(* IEC 61131-3 sources: NachHouse_TST/ROOM_API_PILOT/room_api_pilot, 11 files *)

(* ---- 02_TYPES.ST ---- *)
(*
   ROOM_API_PILOT - d�tov� typy logick�ho API a prenosov�ho protokolu.
   Koment�re opisuj� v�znam pre PLC aj klienta; nejde o re�lnu domov� automatiz�ciu.
*)

TYPE
   NH_API_INFO : STRUCT
    	ApiVersion		: UINT;          (* Verzia verejn�ho API kontraktu. ENG *)
		ApiVarNext		: UINT;          (* Adresa v pam�ti PLC, kde sa nach�dza za�iatok �al��ch premenn�ch API. ENG *)
		ApiVarSize		: UDINT;          (* Ve�kos� v bajtoch, ktor� zaber� v pam�ti PLC. ENG *)
		ApiBussy			: BOOL;          (* TRUE znamen�, �e PLC je zanepr�znene spracovan�m pr�kazu. ENG *)
   END_STRUCT

   NH_LOG_INFO : STRUCT
		BufferBegin		: UDINT;          (* Adresa v pam�ti PLC, kde sa nach�dza za�iatok logovacieho bufferu. ENG *)
		BufferEnd		: UDINT;          (* Adresa v pamti PLC, kde sa nachdza zaiatok logovacieho bufferu. ENG *)
		BufferNext		: UDINT;          (* Adresa v pamti PLC, kde sa nachdza zaiatokalch premennch API. ENG *)
		BufferSize		: UDINT;          (* Vekos v bajtoch, ktor zaber v pamti PLC. ENG *)
   END_STRUCT

END_TYPE

TYPE
    NH_API_DIFF_HEAD : STRUCT                    (* Header pre diff udajov, Sizeof = 40B *)
        StructID        : UINT := 1;          		(* Cislo struktury zaslatych udajov - parser  *)
        Name            : STRING[21] := 'T_ROOM_STATE';   (* What scheme used for parser. StructID = 1 = T_ROOM_STATE*)
        Records         : INT := 2;          		(* Pocet zaslatych zaznamov T_ROOM_STATE *)
        RecSize         : UDINT := 21;      			(* Size of 1. T_ROOM_STATE*)
        MessageSize     : UDINT := 42;      			(* Len Doplnujuce info Records * RecSize := 2*21=42B *)
        HeadIndex       : UINT := 0;						(* index tohto headera ApiVarsPublic[0], koniec ApiVarsPublic[0] + 40B = ApiVarsPublic[3] *)
        BeginIndex      : UINT := 4;          		(* kde zacinaju data struktury = 1.veta ApiVarsPublic[4] *)
        EndIndex        : UINT := 8;          		(* kde koncia data ApiVarsPublic[8] .. len informacne, lebo nemusi byt zaplnenychcelych 4B DWORD *)
	END_STRUCT

	T_ROOM_STATE : STRUCT
      RoomId          : UDINT; (* V?zba stavov?ho z?znamu na stabiln? ID v konfigur?cii. ENG *)
    	Temperature     : REAL;  (* Zobrazovan? testovacia teplota v stup?och Celzia. ENG *)
    	Humidity        : REAL;  (* Zobrazovan? testovacia relat?vna vlhkos? v percent?ch. ENG *)
    	Presence        : BOOL;  (* Testovac? pr?znak pr?tomnosti ovplyv?uj?ci pozadie karty. ENG *)
    	DayPhase        : UINT;  (* K?d dennej f?zy API_DAY_PHASE_* pre existuj?cu ikonu. ENG *)
    	CategoryMask    : DWORD; (* Bitov? maska kateg?ri?, ktor?ch ikony sa maj? zobrazi?. ENG *)
    	AlarmLevel      : USINT; (* Vizu?lna ?rove? API_ALARM_*; nesp???a re?lny alarm. ENG *)
    	Online          : BOOL;  (* Dostupnos? d?t miestnosti pre klienta. ENG *)
	END_STRUCT
END_TYPE
TYPE
   NH_API_DIFF_HEAD : STRUCT                    (* Header pre diff udajov, Sizeof = 40B *)
		StructID		: UINT := 1;          		(* Cislo struktury zaslatych udajov - parser  *)
		Name			: STRING[21] := 'T_ROOM_STATE';   (* What scheme used for parser. StructID = 1 = T_ROOM_STATE*)
		Records			: INT := 2;          		(* Pocet zaslatych zaznamov T_ROOM_STATE *)
		RecSize			: UDINT := 21;      			(* Size of 1. T_ROOM_STATE*)
		MessageSize		: UDINT := 42;      			(* Len Doplnujuce info Records * RecSize := 2*21=42B *)
         HeadIndex      : UINT := 0;						(* index tohto headera ApiVarsPublic[0], koniec ApiVarsPublic[0] + 40B = ApiVarsPublic[3] *)
		BeginIndex		: UINT := 4;          		(* kde zacinaju data struktury = 1.veta ApiVarsPublic[4] *)
		EndIndex		: UINT := 8;          		(* kde koncia data ApiVarsPublic[8] .. len informacne, lebo nemusi byt zaplnenychcelych 4B DWORD *)
	END_STRUCT

	T_ROOM_STATE : STRUCT
   	    RoomId          : UDINT; (* V�zba stavov�ho z�znamu na stabiln� ID v konfigur�cii. ENG *)
    	Temperature     : REAL;  (* Zobrazovan� testovacia teplota v stup�och Celzia. ENG *)
    	Humidity        : REAL;  (* Zobrazovan� testovacia relat�vna vlhkos� v percent�ch. ENG *)
    	Presence        : BOOL;  (* Testovac� pr�znak pr�tomnosti ovplyv�uj�ci pozadie karty. ENG *)
    	DayPhase        : UINT;  (* K�d dennej f�zy API_DAY_PHASE_* pre existuj�cu ikonu. ENG *)
    	CategoryMask    : DWORD; (* Bitov� maska kateg�ri�, ktor�ch ikony sa maj� zobrazi�. ENG *)
    	AlarmLevel      : USINT; (* Vizu�lna �rove� API_ALARM_*; nesp���a re�lny alarm. ENG *)
    	Online          : BOOL;  (* Dostupnos� d�t miestnosti pre klienta. ENG *)
	END_STRUCT
END_TYPE

(* V�sledok vykonania jedn�ho klientsk�ho pr�kazu. *)
TYPE
T_API_COMMAND_RESULT : STRUCT
    ClientId       : STRING[36]; (* Identifik�tor klienta, ktor�mu patr� v�sledok. ENG *)
    RequestId      : UDINT;      (* Identifik�tor po�iadavky pridelen� klientom. ENG *)
    Result         : USINT;      (* ��seln� n�vratov� k�d API_RESULT_*. ENG *)
    Message        : STRING[80]; (* Kr�tky slovensk� text v�sledku ur�en� pre log a testovanie. *)
    ConfigRevision : UDINT;      (* Rev�zia konfigur�cie platn� po spracovan� pr�kazu. ENG *)
    StateRevision  : UDINT;      (* Rev�zia stavov�ch �dajov platn� po spracovan� pr�kazu. ENG *)
END_STRUCT
END_TYPE

(* Z�kladn� inform�cie o API a jeho aktu�lnych rev�zi�ch. *)
TYPE T_API_INFO :
STRUCT
    ApiVersion        : STRING[32];          (* Verzia verejn�ho API kontraktu. ENG *)
    ConfigRevision    : UDINT;               (* Aktu�lna rev�zia konfigur�cie miestnost�. ENG *)
    StateRevision     : UDINT;               (* Aktu�lna rev�zia dynamick�ch stavov miestnost�. ENG *)
    MaxRooms          : USINT;               (* Najvy��� po�et miestnost� podporovan� PLC. ENG *)
    LastCommandResult : T_API_COMMAND_RESULT; (* Posledn� v�sledok pr�kazu, dostupn� aj po obnoven� klienta. ENG *)
END_STRUCT
END_TYPE

(* Konfigura�n� �daje jednej miestnosti. *)
TYPE T_ROOM_CONFIG :
STRUCT
    Used        : BOOL;       (* TRUE znamen�, �e je t�to poz�cia po�a obsaden� miestnos�ou. ENG *)
    RoomId      : UDINT;      (* Stabiln� a jedine�n� identifik�tor miestnosti; hodnota 0 je neplatn�. ENG *)
    Name        : STRING[64]; (* Hlavn� n�zov miestnosti zobrazen� na karte. ENG *)
    ProjectName : STRING[64]; (* Doplnkov� n�zov zobrazen� pod hlavn�m n�zvom. ENG *)
    IconId      : UINT;       (* Identifik�tor ikony pou��vanej frozen browserom. ENG *)
    SortDefault : UINT;       (* Predvolen� poradie iba pri prvom na��tan� klienta. ENG *)
END_STRUCT
END_TYPE

(* �pln� konfigura�n� snapshot v�etk�ch poz�ci� miestnost�. *)
TYPE T_API_CONFIG :
STRUCT
    Rooms : ARRAY[1..40] OF T_ROOM_CONFIG; (* Pevn� pole najviac 40 konfigura�n�ch z�znamov. ENG *)
END_STRUCT
END_TYPE

(* Ru�ne nastavovan� pilotn� stav jednej miestnosti. *)

(* �pln� stavov� snapshot v�etk�ch poz�ci� miestnost�. *)
TYPE T_API_STATE :
STRUCT
    Rooms : ARRAY[1..40] OF T_ROOM_STATE; (* Pevn� pole najviac 40 stavov�ch z�znamov. ENG *)
END_STRUCT
END_TYPE

(* Po�iadavka klienta na pridanie, zmazanie, kop�rovanie alebo �pravu miestnosti. *)
TYPE T_API_COMMAND_ROOM :
STRUCT
    ClientId     : STRING[36]; (* Identifik�tor klienta odosielaj�ceho pr�kaz. ENG *)
    RequestId    : UDINT;      (* Nenulov� identifik�tor po�iadavky pre p�rovanie a opakovanie. ENG *)
    Action       : USINT;      (* Po�adovan� akcia ur�en� kon�tantou API_ACTION_*. ENG *)
    RoomId       : UDINT;      (* Cie�ov� stabiln� ID miestnosti. ENG *)
    SourceRoomId : UDINT;      (* Zdrojov� ID pou�it� iba pri kop�rovan� miestnosti. ENG *)
    Name         : STRING[64]; (* Nov� alebo upraven� hlavn� n�zov miestnosti. ENG *)
    ProjectName  : STRING[64]; (* Nov� alebo upraven� doplnkov� n�zov miestnosti. ENG *)
END_STRUCT
END_TYPE

(* Jedna polo�ka konfigura�n�ho diffu. *)
TYPE T_API_CONFIG_CHANGE :
STRUCT
    Valid     : BOOL;          (* TRUE znamen�, �e polo�ka obsahuje platn� zmenu. ENG *)
    Operation : USINT;         (* Druh zmeny API_DIFF_UPSERT alebo API_DIFF_DELETE. ENG *)
    RoomId    : UDINT;         (* Stabiln� ID zmenenej alebo odstr�nenej miestnosti. ENG *)
    Room      : T_ROOM_CONFIG; (* �pln� nov� z�znam pri UPSERT; pri DELETE je vy�isten�. ENG *)
END_STRUCT
END_TYPE

(* Jedna polo�ka stavov�ho diffu. *)
TYPE T_API_STATE_CHANGE :
STRUCT
    Valid     : BOOL;         (* TRUE znamen�, �e polo�ka obsahuje platn� zmenu. ENG *)
    Operation : USINT;        (* Druh zmeny API_DIFF_UPSERT alebo API_DIFF_DELETE. ENG *)
    RoomId    : UDINT;        (* Stabiln� ID zmenen�ho alebo odstr�nen�ho stavu. ENG *)
    Room      : T_ROOM_STATE; (* �pln� nov� stav pri UPSERT; pri DELETE je vy�isten�. ENG *)
END_STRUCT
END_TYPE

(* Jeden rev�zny r�mec zmien konfigur�cie. *)
TYPE T_API_CONFIG_DIFF :
STRUCT
    Valid        : BOOL;  (* TRUE znamen�, �e hlavi�ka a obsah r�mca s� pripraven�. ENG *)
    FromRevision : UDINT; (* Rev�zia, na ktor� tento r�mec priamo nadv�zuje. ENG *)
    ToRevision   : UDINT; (* Rev�zia po aplikovan� v�etk�ch zmien z r�mca. ENG *)
    FullRequired : BOOL;  (* TRUE prikazuje klientovi na��ta� cel� snapshot. ENG *)
    ChangeCount  : USINT; (* Po�et platn�ch polo�iek na za�iatku po�a Changes. ENG *)
    Changes      : ARRAY[1..40] OF T_API_CONFIG_CHANGE; (* Zmeny konfigur�cie patriace do jednej rev�zie. ENG *)
END_STRUCT
END_TYPE

(* Jeden rev�zny r�mec zmien dynamick�ho stavu. *)
TYPE T_API_STATE_DIFF :
STRUCT
    Valid        : BOOL;  (* TRUE znamen�, �e hlavi�ka a obsah r�mca s� pripraven�. ENG *)
    FromRevision : UDINT; (* Rev�zia, na ktor� tento r�mec priamo nadv�zuje. ENG *)
    ToRevision   : UDINT; (* Rev�zia po aplikovan� v�etk�ch zmien z r�mca. ENG *)
    FullRequired : BOOL;  (* TRUE prikazuje klientovi na��ta� cel� snapshot. ENG *)
    ChangeCount  : USINT; (* Po�et platn�ch polo�iek na za�iatku po�a Changes. ENG *)
    Changes      : ARRAY[1..40] OF T_API_STATE_CHANGE; (* Stavov� zmeny patriace do jednej rev�zie. ENG *)
END_STRUCT
END_TYPE

(* Po�iadavka transportn�ho handshake na z�skanie �al�ieho uchovan�ho diffu. ENG *)
TYPE T_API_SYNC_REQUEST :
STRUCT
    ClientId           : STRING[36]; (* Identifik�tor klienta �iadaj�ceho synchroniz�ciu. ENG *)
    RequestId          : UDINT;      (* Nenulov� identifik�tor synchroniza�nej po�iadavky. ENG *)
    ConfigFromRevision : UDINT;      (* Posledn� konfigura�n� rev�zia �spe�ne ulo�en� klientom. ENG *)
    StateFromRevision  : UDINT;      (* Posledn� stavov� rev�zia �spe�ne ulo�en� klientom. ENG *)
END_STRUCT
END_TYPE

(* Odpove� PLC na jednu synchroniza�n� po�iadavku. *)
TYPE T_API_SYNC_RESPONSE :
STRUCT
    ClientId   : STRING[36];       (* Identifik�tor klienta prevzat� z po�iadavky. ENG *)
    RequestId  : UDINT;            (* Identifik�tor po�iadavky prevzat� z po�iadavky. ENG *)
    Result     : USINT;            (* Celkov� n�vratov� k�d synchroniz�cie API_RESULT_*. ENG *)
    Message    : STRING[80];       (* Kr�tky slovensk� opis v�sledku pre log a testovanie. *)
    ConfigMode : USINT;            (* Re�im konfigura�nej odpovede API_SYNC_*. ENG *)
    StateMode  : USINT;            (* Re�im stavovej odpovede API_SYNC_*. ENG *)
    ConfigDiff : T_API_CONFIG_DIFF; (* �al�� konfigura�n� r�mec alebo po�iadavka na cel� snapshot. ENG *)
    StateDiff  : T_API_STATE_DIFF; (* �al�� stavov� r�mec alebo po�iadavka na cel� snapshot. ENG *)
END_STRUCT
END_TYPE

(* Ru�n� testovac� vstup oddelen� od produk�n�ho pr�kazu ApiCommandRoom. *)
TYPE T_API_TEST_STATE_REQUEST :
STRUCT
    ClientId     : STRING[36]; (* Identifik�tor testovacieho klienta. ENG *)
    RequestId    : UDINT;      (* Nenulov� identifik�tor testovacej po�iadavky. ENG *)
    RoomId       : UDINT;      (* Stabiln� ID miestnosti, ktorej stav sa m� zmeni�. ENG *)
    Temperature  : REAL;       (* Po�adovan� testovacia teplota od -50 do 100 �C. ENG *)
    Humidity     : REAL;       (* Po�adovan� testovacia vlhkos� od 0 do 100 %. ENG *)
    Presence     : BOOL;       (* Po�adovan� testovac� pr�znak pr�tomnosti. ENG *)
    DayPhase     : UINT;       (* Po�adovan� platn� denn� f�za API_DAY_PHASE_*. ENG *)
    CategoryMask : DWORD;      (* Po�adovan� bitov� maska kateg�ri�. ENG *)
    AlarmLevel   : USINT;      (* Po�adovan� vizu�lna �rove� API_ALARM_*. ENG *)
    Online       : BOOL;       (* Po�adovan� testovacia dostupnos� d�t. ENG *)
END_STRUCT
END_TYPE

(* ---- 01_CONSTANTS.ST ---- *)
(*
   ROOM_API_PILOT - verejn� ��seln� kontrakt a pevn� limity pilotu.
   ��seln� hodnoty s� s��as�ou API; klient ich nesmie svojvo�ne meni�.
*)

VAR_GLOBAL CONSTANT
    C_API_VERSION          : STRING[32] := 'ROOM_API_PILOT/1'; (* Textov� verzia verejn�ho API kontraktu. ENG *)
    C_MAX_ROOMS            : USINT := 40;                     (* Najvy��� po�et miestnost� podporovan� pilotom. *)
    C_DIFF_HISTORY_DEPTH   : USINT := 8;                      (* Po�et uchov�van�ch r�mcov zmien v kruhovej hist�rii. *)

    (* ��seln� k�dy akci� po�a Action v pr�kaze miestnosti. *)
    API_ACTION_NONE          : USINT := 0; (* Nie je zvolen� �iadna akcia. ENG *)
    API_ACTION_ADD_ROOM      : USINT := 1; (* Pridanie novej miestnosti. ENG *)
    API_ACTION_DELETE_ROOM   : USINT := 2; (* Odstr�nenie existuj�cej miestnosti. ENG *)
    API_ACTION_COPY_ROOM     : USINT := 3; (* Vytvorenie k�pie existuj�cej miestnosti. ENG *)
    API_ACTION_SET_ROOM_DATA : USINT := 4; (* Zmena n�zvov�ch �dajov miestnosti. ENG *)

    (* ��seln� n�vratov� k�dy po�a Result. *)
    API_RESULT_NONE               : USINT := 0; (* V�sledok e�te nie je k dispoz�cii. ENG *)
    API_RESULT_OK                 : USINT := 1; (* Oper�cia prebehla �spe�ne. ENG *)
    API_RESULT_ERROR              : USINT := 2; (* V�eobecn�, bli��ie neur�en� chyba. ENG *)
    API_RESULT_NOT_FOUND          : USINT := 3; (* Po�adovan� objekt sa nena�iel. ENG *)
    API_RESULT_NO_FREE_SLOT       : USINT := 4; (* Nie je vo�n� poz�cia pre �al�iu miestnos�. ENG *)
    API_RESULT_ALREADY_EXISTS     : USINT := 5; (* Objekt s rovnak�m identifik�torom u� existuje. ENG *)
    API_RESULT_INVALID_ARGUMENT   : USINT := 6; (* Aspo� jeden vstupn� �daj je neplatn�. ENG *)
    API_RESULT_UNSUPPORTED_ACTION : USINT := 7; (* Klient po�aduje nepodporovan� akciu. ENG *)

    (* Druh oper�cie zap�sanej v jednom z�zname diffu. *)
    API_DIFF_NONE   : USINT := 0; (* Z�znam neobsahuje zmenu. ENG *)
    API_DIFF_UPSERT : USINT := 1; (* Vlo�enie nov�ho alebo �pln� aktualiz�cia existuj�ceho z�znamu. ENG *)
    API_DIFF_DELETE : USINT := 2; (* Odstr�nenie z�znamu. ENG *)

    (* Re�im odpovede synchroniza�n�ho mechanizmu. *)
    API_SYNC_CURRENT       : USINT := 0; (* Cache klienta u� zodpoved� aktu�lnej rev�zii. ENG *)
    API_SYNC_DIFF          : USINT := 1; (* Odpove� obsahuje jeden nadv�zuj�ci r�mec zmien. ENG *)
    API_SYNC_FULL_REQUIRED : USINT := 2; (* Hist�ria nesta�� a klient mus� na��ta� cel� snapshot. ENG *)

    (* Vizu�lna �rove� alarmu zobrazovan� na karte miestnosti. *)
    API_ALARM_OK      : USINT := 0; (* Bez upozornenia alebo alarmu. ENG *)
    API_ALARM_WARNING : USINT := 1; (* Upozornenie. ENG *)
    API_ALARM_ALARM   : USINT := 2; (* Alarm. ENG *)

    (* Identifik�tory existuj�cich ikon dennej f�zy vo frozen browseri V0.5.72. *)
    API_DAY_PHASE_DAY   : UINT := 140; (* Denn� f�za. ENG *)
    API_DAY_PHASE_DUSK  : UINT := 142; (* S�mrak. ENG *)
    API_DAY_PHASE_NIGHT : UINT := 144; (* No�n� f�za. ENG *)
    API_DAY_PHASE_DAWN  : UINT := 146; (* �svit. ENG *)

    (* Predvolen� testovacie hodnoty pou�it� pri pridan� miestnosti. *)
    API_DEFAULT_ICON_ID     : UINT := 16;   (* Predvolen� identifik�tor ikony miestnosti. *)
    API_DEFAULT_TEMPERATURE : REAL := 20.0; (* Predvolen� teplota v stup�och Celzia. *)
    API_DEFAULT_HUMIDITY    : REAL := 40.0; (* Predvolen� relat�vna vlhkos� v percent�ch. *)
END_VAR

(* ---- 03_PUBLIC_API.ST ---- *)
(*
   V�etky objekty vidite�n� klientom s� glob�lne a ozna�en� atrib�tom PUBLIC_API.
   Klient mus� najprv zap�sa� cel� obsah po�iadavky a pr�znak Execute a� ako posledn�.
   Snapshoty ApiConfig a ApiState s� pod�a kontraktu ur�en� iba na ��tanie.
   N�zvy verejn�ch objektov tvoria stabiln� anglick� API kontrakt. ENG
*)

VAR_GLOBAL
    ApiInfo       {PUBLIC_API} : T_API_INFO;   (* Inform�cie o verzii, rev�zi�ch, limite a poslednom pr�kaze. ENG *)
    ApiConfig     {PUBLIC_API} : T_API_CONFIG; (* �pln� konfigura�n� snapshot ur�en� klientovi iba na ��tanie. ENG *)
    ApiState      {PUBLIC_API} : T_API_STATE;  (* �pln� stavov� snapshot ur�en� klientovi iba na ��tanie. ENG *)

    ApiConfigDiff {PUBLIC_API} : T_API_CONFIG_DIFF; (* Najnov�� vytvoren� r�mec zmien konfigur�cie. ENG *)
    ApiStateDiff  {PUBLIC_API} : T_API_STATE_DIFF;  (* Najnov�� vytvoren� r�mec zmien stavu. ENG *)

    (* Dvojf�zov� kan�l pr�kazov miestnosti: payload, Execute, spracovanie, Finished. ENG *)
    ApiCommandRoom     {PUBLIC_API} : T_API_COMMAND_ROOM;  (* Obsah po�iadavky zapisovan� klientom. ENG *)
    ApiCommandExecute  {PUBLIC_API} : BOOL;                (* Sp���ac� pr�znak; klient ho zapisuje ako posledn�. ENG *)
    ApiCommandBusy     {PUBLIC_API} : BOOL;                (* TRUE po�as spracovania pr�kazu v PLC. ENG *)
    ApiCommandFinished {PUBLIC_API} : BOOL;                (* TRUE po dokon�en�; klient m��e pre��ta� v�sledok. ENG *)
    ApiCommandResult   {PUBLIC_API} : T_API_COMMAND_RESULT; (* V�sledok pr�ve dokon�en�ho alebo zopakovan�ho pr�kazu. ENG *)

    (* Dvojf�zov� kan�l obnovy cache a na��tania jedn�ho nadv�zuj�ceho diffu. ENG *)
    ApiSyncRequest  {PUBLIC_API} : T_API_SYNC_REQUEST;  (* Rev�zie, od ktor�ch chce klient pokra�ova�. ENG *)
    ApiSyncExecute  {PUBLIC_API} : BOOL;                (* Sp���ac� pr�znak synchroniz�cie zapisovan� ako posledn�. ENG *)
    ApiSyncBusy     {PUBLIC_API} : BOOL;                (* TRUE po�as pr�pravy synchroniza�nej odpovede. ENG *)
    ApiSyncFinished {PUBLIC_API} : BOOL;                (* TRUE po pripraven� odpovede pre klienta. ENG *)
    ApiSyncResponse {PUBLIC_API} : T_API_SYNC_RESPONSE; (* V�sledn� re�imy a najviac jeden diff ka�dej vetvy. ENG *)

    (* Samostatn� kan�l ru�n�ho nastavovania pilotn�ch stavov bez re�lneho IO. *)
    ApiTestStateRequest  {PUBLIC_API} : T_API_TEST_STATE_REQUEST; (* Testovacie stavov� hodnoty zapisovan� klientom. ENG *)
    ApiTestStateExecute  {PUBLIC_API} : BOOL;                     (* Sp���ac� pr�znak testovacieho z�pisu. ENG *)
    ApiTestStateBusy     {PUBLIC_API} : BOOL;                     (* TRUE po�as valid�cie a z�pisu testovacieho stavu. ENG *)
    ApiTestStateFinished {PUBLIC_API} : BOOL;                     (* TRUE po dokon�en� testovacieho z�pisu. ENG *)
    ApiTestStateResult   {PUBLIC_API} : T_API_COMMAND_RESULT;     (* V�sledok posledn�ho testovacieho z�pisu. ENG *)

	ApiVarsPublic 	{PUBLIC_API} : ARRAY[0..999] OF DWORD; (* Jedina komunikacna oblast binarnychch Vars, ktoru naplna PLC zmenami*)

	SizeApiHeder 	: UDINT;
	SizeStructRoom	: UDINT;
	SizeApiVars	: UDINT;

	Ptr_T_ROOM_STATE_Src    : PTR_TO T_ROOM_STATE;
   Ptr_T_ROOM_STATE_Dest   : PTR_TO T_ROOM_STATE;

END_VAR

(* ---- 04_INTERNAL.ST ---- *)
(*
   Interné pracovné údaje PLC sa neexportujú do TecoApi ani PLCComS.
   Klient k nim nemá pristupovať a nie sú súčasťou verejného kontraktu.
*)

VAR_GLOBAL
    ApiInitialized : BOOL; (* TRUE po jednorazovom dokončení inicializácie pilotných dát. ENG *)

    (* Tieňové kópie posledného zachyteného snapshotu používané na výpočet zmien. *)
    ApiConfigShadow : ARRAY[1..40] OF T_ROOM_CONFIG; (* Posledná známa konfigurácia pre porovnanie. ENG *)
    ApiStateShadow  : ARRAY[1..40] OF T_ROOM_STATE;  (* Posledný známy stav pre porovnanie. ENG *)

    (* Kruhové histórie ôsmich posledných revíznych rámcov pre obnovu cache klienta. *)
    ApiConfigDiffHistory : ARRAY[1..8] OF T_API_CONFIG_DIFF; (* Uchované konfiguračné diffy. ENG *)
    ApiStateDiffHistory  : ARRAY[1..8] OF T_API_STATE_DIFF;  (* Uchované stavové diffy. ENG *)
    ApiConfigHistoryHead : USINT; (* Index najnovšieho konfiguračného rámca; 0 pred prvým zápisom. ENG *)
    ApiStateHistoryHead  : USINT; (* Index najnovšieho stavového rámca; 0 pred prvým zápisom. ENG *)

    (* Údaje potrebné na idempotentné zopakovanie bezprostredne posledného príkazu. *)
    ApiLastCommandClientId  : STRING[36];          (* ClientId posledného spracovaného príkazu. ENG *)
    ApiLastCommandRequestId : UDINT;               (* RequestId posledného spracovaného príkazu. ENG *)
    ApiLastStoredResult     : T_API_COMMAND_RESULT; (* Úplný uložený výsledok posledného príkazu. ENG *)
END_VAR

(* ---- 05_UTILS.ST ---- *)
(* ROOM_API_PILOT - malé deterministické pomocné funkcie bez skrytého stavu. *)

(* Porovná všetky polia dvoch konfiguračných záznamov miestnosti. *)
FUNCTION ApiRoomConfigEqual : BOOL
VAR_INPUT
    A : T_ROOM_CONFIG; (* Prvý porovnávaný konfiguračný záznam. *)
    B : T_ROOM_CONFIG; (* Druhý porovnávaný konfiguračný záznam. *)
END_VAR

(* TRUE sa vráti iba vtedy, keď sú všetky polia zhodné. *)
ApiRoomConfigEqual :=
    (A.Used = B.Used) AND
    (A.RoomId = B.RoomId) AND
    (A.Name = B.Name) AND
    (A.ProjectName = B.ProjectName) AND
    (A.IconId = B.IconId) AND
    (A.SortDefault = B.SortDefault);
END_FUNCTION

(* Porovná všetky polia dvoch stavových záznamov miestnosti. *)
FUNCTION ApiRoomStateEqual : BOOL
VAR_INPUT
    A : T_ROOM_STATE; (* Prvý porovnávaný stavový záznam. *)
    B : T_ROOM_STATE; (* Druhý porovnávaný stavový záznam. *)
END_VAR

(* TRUE sa vráti iba vtedy, keď sú všetky polia zhodné. *)
ApiRoomStateEqual :=
    (A.RoomId = B.RoomId) AND
    (A.Temperature = B.Temperature) AND
    (A.Humidity = B.Humidity) AND
    (A.Presence = B.Presence) AND
    (A.DayPhase = B.DayPhase) AND
    (A.CategoryMask = B.CategoryMask) AND
    (A.AlarmLevel = B.AlarmLevel) AND
    (A.Online = B.Online);
END_FUNCTION

(* Vyhľadá obsadenú konfiguračnú pozíciu podľa stabilného RoomId. *)
FUNCTION ApiFindConfigSlot : USINT
VAR_INPUT
    RoomId : UDINT; (* Hľadané stabilné ID; hodnota 0 sa zámerne nehľadá. ENG *)
END_VAR
VAR
    i : USINT; (* Index pre prechod poľom miestností. *)
END_VAR

(* Hodnota 0 znamená, že miestnosť nebola nájdená. *)
ApiFindConfigSlot := 0;
IF RoomId <> 0 THEN
    FOR i := 1 TO C_MAX_ROOMS DO
        IF ApiConfig.Rooms[i].Used AND (ApiConfig.Rooms[i].RoomId = RoomId) THEN
            ApiFindConfigSlot := i;
            RETURN;
        END_IF;
    END_FOR;
END_IF;
END_FUNCTION

(* Vyhľadá stavovú pozíciu podľa stabilného RoomId. *)
FUNCTION ApiFindStateSlot : USINT
VAR_INPUT
    RoomId : UDINT; (* Hľadané stabilné ID; hodnota 0 sa zámerne nehľadá. ENG *)
END_VAR
VAR
    i : USINT; (* Index pre prechod poľom stavov. *)
END_VAR

(* Hodnota 0 znamená, že stav miestnosti nebol nájdený. *)
ApiFindStateSlot := 0;
IF RoomId <> 0 THEN
    FOR i := 1 TO C_MAX_ROOMS DO
        IF ApiState.Rooms[i].RoomId = RoomId THEN
            ApiFindStateSlot := i;
            RETURN;
        END_IF;
    END_FOR;
END_IF;
END_FUNCTION

(* Nájde prvú voľnú pozíciu v konfiguračnom poli. *)
FUNCTION ApiFindFreeConfigSlot : USINT
VAR
    i : USINT; (* Index pre prechod poľom miestností. *)
END_VAR

(* Hodnota 0 znamená, že všetkých 40 pozícií je obsadených. *)
ApiFindFreeConfigSlot := 0;
FOR i := 1 TO C_MAX_ROOMS DO
    IF NOT ApiConfig.Rooms[i].Used THEN
        ApiFindFreeConfigSlot := i;
        RETURN;
    END_IF;
END_FOR;
END_FUNCTION

(* Nájde prvú voľnú pozíciu v stavovom poli. *)
FUNCTION ApiFindFreeStateSlot : USINT
VAR
    i : USINT; (* Index pre prechod poľom stavov. *)
END_VAR

(* Voľný stavový slot je označený hodnotou RoomId = 0. ENG *)
ApiFindFreeStateSlot := 0;
FOR i := 1 TO C_MAX_ROOMS DO
    IF ApiState.Rooms[i].RoomId = 0 THEN
        ApiFindFreeStateSlot := i;
        RETURN;
    END_IF;
END_FOR;
END_FUNCTION

(* Vynuluje konfiguračný záznam a označí jeho pozíciu ako nepoužitú. *)
FUNCTION ApiClearRoomConfig : BOOL
VAR_IN_OUT
    Room : T_ROOM_CONFIG; (* Konfiguračný záznam odovzdaný referenciou na vyčistenie. *)
END_VAR

(* Každé pole sa nastavuje explicitne kvôli deterministickému výsledku. *)
Room.Used := FALSE;
Room.RoomId := 0;
Room.Name := '';
Room.ProjectName := '';
Room.IconId := 0;
Room.SortDefault := 0;
ApiClearRoomConfig := TRUE;
END_FUNCTION

(* Vynuluje stavový záznam a uvoľní jeho pozíciu hodnotou RoomId = 0. *)
FUNCTION ApiClearRoomState : BOOL
VAR_IN_OUT
    Room : T_ROOM_STATE; (* Stavový záznam odovzdaný referenciou na vyčistenie. *)
END_VAR

(* Bezpečné nulové hodnoty nepredstavujú žiadnu reálnu IO informáciu. *)
Room.RoomId := 0;
Room.Temperature := 0.0;
Room.Humidity := 0.0;
Room.Presence := FALSE;
Room.DayPhase := API_DAY_PHASE_DAY;
Room.CategoryMask := DWORD#16#00000000;
Room.AlarmLevel := API_ALARM_OK;
Room.Online := FALSE;
ApiClearRoomState := TRUE;
END_FUNCTION

(* Vyčistí hlavičku aj všetkých 40 položiek konfiguračného diffu. *)
FUNCTION ApiClearConfigDiff : BOOL
VAR_IN_OUT
    Diff : T_API_CONFIG_DIFF; (* Konfiguračný rámec odovzdaný referenciou na vyčistenie. ENG *)
END_VAR
VAR
    i : USINT; (* Index pre vyčistenie celého poľa Changes. ENG *)
END_VAR

(* Po vyčistení rámec nie je platný, kým ho producent znova nenaplní. *)
Diff.Valid := FALSE;
Diff.FromRevision := 0;
Diff.ToRevision := 0;
Diff.FullRequired := FALSE;
Diff.ChangeCount := 0;
FOR i := 1 TO C_MAX_ROOMS DO
    Diff.Changes[i].Valid := FALSE;
    Diff.Changes[i].Operation := API_DIFF_NONE;
    Diff.Changes[i].RoomId := 0;
    ApiClearRoomConfig(Diff.Changes[i].Room);
END_FOR;
ApiClearConfigDiff := TRUE;
END_FUNCTION

(* Vyčistí hlavičku aj všetkých 40 položiek stavového diffu. *)
FUNCTION ApiClearStateDiff : BOOL
VAR_IN_OUT
    Diff : T_API_STATE_DIFF; (* Stavový rámec odovzdaný referenciou na vyčistenie. ENG *)
END_VAR
VAR
    i : USINT; (* Index pre vyčistenie celého poľa Changes. ENG *)
END_VAR

(* Po vyčistení rámec nie je platný, kým ho producent znova nenaplní. *)
Diff.Valid := FALSE;
Diff.FromRevision := 0;
Diff.ToRevision := 0;
Diff.FullRequired := FALSE;
Diff.ChangeCount := 0;
FOR i := 1 TO C_MAX_ROOMS DO
    Diff.Changes[i].Valid := FALSE;
    Diff.Changes[i].Operation := API_DIFF_NONE;
    Diff.Changes[i].RoomId := 0;
    ApiClearRoomState(Diff.Changes[i].Room);
END_FOR;
ApiClearStateDiff := TRUE;
END_FUNCTION

(* Vypočíta nasledujúcu nenulovú revíziu s ošetrením pretečenia UDINT. *)
FUNCTION ApiNextRevision : UDINT
VAR_INPUT
    Revision : UDINT; (* Aktuálna revízia, z ktorej sa má vytvoriť nasledovník. ENG *)
END_VAR

ApiNextRevision := Revision + 1;
(* Hodnota 0 je vyhradená pre klienta bez načítaného snapshotu. *)
IF ApiNextRevision = 0 THEN
    ApiNextRevision := 1;
END_IF;
END_FUNCTION

(* Overí, či hodnota patrí medzi štyri denné fázy podporované browserom. *)
FUNCTION ApiValidDayPhase : BOOL
VAR_INPUT
    DayPhase : UINT; (* Kontrolovaný identifikátor dennej fázy. ENG *)
END_VAR

ApiValidDayPhase :=
    (DayPhase = API_DAY_PHASE_DAY) OR
    (DayPhase = API_DAY_PHASE_DUSK) OR
    (DayPhase = API_DAY_PHASE_NIGHT) OR
    (DayPhase = API_DAY_PHASE_DAWN);
END_FUNCTION

(* ---- 06_DIFF_ENGINE.ST ---- *)
(*
   Mechanizmus výpočtu rozdielov (diff engine). ENG
   Jedna PLC transakcia vytvorí jednu novú revíziu a jeden úplný rámec zmien.
   Uchováva sa osem rámcov; klient si vyžiada vždy práve jeden nasledujúci rámec.
*)

(* Zachytí všetky konfiguračné zmeny od poslednej tieňovej kópie. *)
FUNCTION ApiCaptureConfigChanges : BOOL
VAR
    i          : USINT; (* Index pri prechode všetkých konfiguračných pozícií. *)
    count      : USINT; (* Počet zmien zapísaných do aktuálneho rámca. ENG *)
    oldRev     : UDINT; (* Revízia konfigurácie pred zachytením zmien. ENG *)
    newRev     : UDINT; (* Nová revízia konfigurácie po zachytení zmien. ENG *)
    anyChanged : BOOL;  (* Pomocný príznak, že sa zmenila aspoň jedna pozícia. ENG *)
END_VAR

(* Prvý prechod iba zisťuje, či treba vytvoriť novú revíziu. *)
anyChanged := FALSE;
FOR i := 1 TO C_MAX_ROOMS DO
    IF NOT ApiRoomConfigEqual(ApiConfig.Rooms[i], ApiConfigShadow[i]) THEN
        anyChanged := TRUE;
    END_IF;
END_FOR;

ApiCaptureConfigChanges := anyChanged;
(* Bez zmeny sa revízia ani história neposúvajú. *)
IF NOT anyChanged THEN
    RETURN;
END_IF;

(* Pripraví hlavičku nového konfiguračného rámca. *)
ApiClearConfigDiff(ApiConfigDiff);
oldRev := ApiInfo.ConfigRevision;
newRev := ApiNextRevision(oldRev);
ApiConfigDiff.FromRevision := oldRev;
ApiConfigDiff.ToRevision := newRev;
ApiConfigDiff.FullRequired := FALSE;
count := 0;

(* Druhý prechod vytvorí kompaktný zoznam UPSERT/DELETE zmien. ENG *)
FOR i := 1 TO C_MAX_ROOMS DO
    IF NOT ApiRoomConfigEqual(ApiConfig.Rooms[i], ApiConfigShadow[i]) THEN
        count := count + 1;
        ApiConfigDiff.Changes[count].Valid := TRUE;

        IF ApiConfig.Rooms[i].Used THEN
            ApiConfigDiff.Changes[count].Operation := API_DIFF_UPSERT;
            ApiConfigDiff.Changes[count].RoomId := ApiConfig.Rooms[i].RoomId;
            ApiConfigDiff.Changes[count].Room := ApiConfig.Rooms[i];
        ELSE
            ApiConfigDiff.Changes[count].Operation := API_DIFF_DELETE;
            ApiConfigDiff.Changes[count].RoomId := ApiConfigShadow[i].RoomId;
            ApiClearRoomConfig(ApiConfigDiff.Changes[count].Room);
        END_IF;
    END_IF;

    ApiConfigShadow[i] := ApiConfig.Rooms[i];
END_FOR;

(* Zverejnenie rámca a revízie sa vykoná až po naplnení všetkých položiek. *)
ApiConfigDiff.ChangeCount := count;
ApiConfigDiff.Valid := TRUE;
ApiInfo.ConfigRevision := newRev;

(* Uloženie hotového rámca do osemprvkovej kruhovej histórie. *)
IF ApiConfigHistoryHead >= C_DIFF_HISTORY_DEPTH THEN
    ApiConfigHistoryHead := 1;
ELSE
    ApiConfigHistoryHead := ApiConfigHistoryHead + 1;
END_IF;
ApiConfigDiffHistory[ApiConfigHistoryHead] := ApiConfigDiff;
END_FUNCTION

(* Zachytí všetky stavové zmeny od poslednej tieňovej kópie. *)
FUNCTION ApiCaptureStateChanges : BOOL
VAR
    i          : USINT; (* Index pri prechode všetkých stavových pozícií. *)
    count      : USINT; (* Počet zmien zapísaných do aktuálneho rámca. ENG *)
    oldRev     : UDINT; (* Revízia stavu pred zachytením zmien. ENG *)
    newRev     : UDINT; (* Nová revízia stavu po zachytení zmien. ENG *)
    anyChanged : BOOL;  (* Pomocný príznak, že sa zmenila aspoň jedna pozícia. ENG *)
END_VAR

(* Prvý prechod iba zisťuje, či treba vytvoriť novú revíziu. *)
anyChanged := FALSE;
FOR i := 1 TO C_MAX_ROOMS DO
    IF NOT ApiRoomStateEqual(ApiState.Rooms[i], ApiStateShadow[i]) THEN
        anyChanged := TRUE;
    END_IF;
END_FOR;

ApiCaptureStateChanges := anyChanged;
(* Bez zmeny sa revízia ani história neposúvajú. *)
IF NOT anyChanged THEN
    RETURN;
END_IF;

(* Pripraví hlavičku nového stavového rámca. *)
ApiClearStateDiff(ApiStateDiff);
oldRev := ApiInfo.StateRevision;
newRev := ApiNextRevision(oldRev);
ApiStateDiff.FromRevision := oldRev;
ApiStateDiff.ToRevision := newRev;
ApiStateDiff.FullRequired := FALSE;
count := 0;

(* Druhý prechod vytvorí kompaktný zoznam UPSERT/DELETE zmien. ENG *)
FOR i := 1 TO C_MAX_ROOMS DO
    IF NOT ApiRoomStateEqual(ApiState.Rooms[i], ApiStateShadow[i]) THEN
        count := count + 1;
        ApiStateDiff.Changes[count].Valid := TRUE;

        IF ApiState.Rooms[i].RoomId <> 0 THEN
            ApiStateDiff.Changes[count].Operation := API_DIFF_UPSERT;
            ApiStateDiff.Changes[count].RoomId := ApiState.Rooms[i].RoomId;
            ApiStateDiff.Changes[count].Room := ApiState.Rooms[i];
        ELSE
            ApiStateDiff.Changes[count].Operation := API_DIFF_DELETE;
            ApiStateDiff.Changes[count].RoomId := ApiStateShadow[i].RoomId;
            ApiClearRoomState(ApiStateDiff.Changes[count].Room);
        END_IF;
    END_IF;

    ApiStateShadow[i] := ApiState.Rooms[i];
END_FOR;

(* Zverejnenie rámca a revízie sa vykoná až po naplnení všetkých položiek. *)
ApiStateDiff.ChangeCount := count;
ApiStateDiff.Valid := TRUE;
ApiInfo.StateRevision := newRev;

(* Uloženie hotového rámca do osemprvkovej kruhovej histórie. *)
IF ApiStateHistoryHead >= C_DIFF_HISTORY_DEPTH THEN
    ApiStateHistoryHead := 1;
ELSE
    ApiStateHistoryHead := ApiStateHistoryHead + 1;
END_IF;
ApiStateDiffHistory[ApiStateHistoryHead] := ApiStateDiff;
END_FUNCTION

(* ---- 07_INIT.ST ---- *)
(* Inicializácia pri studenom štarte a deterministické dáta ROOM_API_PILOT. *)

(* Jednorazovo pripraví všetky verejné aj interné objekty pilotu. *)
FUNCTION ApiPilotInit : BOOL
VAR
    i : USINT; (* Index pri inicializácii pevných polí a histórií. *)
END_VAR

(* Opakované volanie po inicializácii už nijaké dáta nemení. *)
ApiPilotInit := ApiInitialized;
IF ApiInitialized THEN
    RETURN;
END_IF;

(* Najprv sa deterministicky vyčistia snapshoty aj ich tieňové kópie. *)
FOR i := 1 TO C_MAX_ROOMS DO
    ApiClearRoomConfig(ApiConfig.Rooms[i]);
    ApiClearRoomState(ApiState.Rooms[i]);
    ApiClearRoomConfig(ApiConfigShadow[i]);
    ApiClearRoomState(ApiStateShadow[i]);
END_FOR;

(* Vyčistenie všetkých pozícií oboch kruhových histórií diffov. ENG *)
FOR i := 1 TO C_DIFF_HISTORY_DEPTH DO
    ApiClearConfigDiff(ApiConfigDiffHistory[i]);
    ApiClearStateDiff(ApiStateDiffHistory[i]);
END_FOR;

(* Štyri ukážkové konfigurácie; všetky hodnoty sú iba testovacie dáta. *)
(* Miestnosť 1: obývačka. *)
ApiConfig.Rooms[1].Used := TRUE;
ApiConfig.Rooms[1].RoomId := 1;
ApiConfig.Rooms[1].Name := 'Obyvacka';
ApiConfig.Rooms[1].ProjectName := '1.01';
ApiConfig.Rooms[1].IconId := 16;
ApiConfig.Rooms[1].SortDefault := 1;

(* Miestnosť 2: kuchyňa. *)
ApiConfig.Rooms[2].Used := TRUE;
ApiConfig.Rooms[2].RoomId := 2;
ApiConfig.Rooms[2].Name := 'Kuchyna';
ApiConfig.Rooms[2].ProjectName := '1.07';
ApiConfig.Rooms[2].IconId := 16;
ApiConfig.Rooms[2].SortDefault := 2;

(* Miestnosť 3: spálňa. *)
ApiConfig.Rooms[3].Used := TRUE;
ApiConfig.Rooms[3].RoomId := 3;
ApiConfig.Rooms[3].Name := 'Spalna';
ApiConfig.Rooms[3].ProjectName := '1.09';
ApiConfig.Rooms[3].IconId := 16;
ApiConfig.Rooms[3].SortDefault := 3;

(* Miestnosť 4: terasa. *)
ApiConfig.Rooms[4].Used := TRUE;
ApiConfig.Rooms[4].RoomId := 4;
ApiConfig.Rooms[4].Name := 'Terasa';
ApiConfig.Rooms[4].ProjectName := 'E.01';
ApiConfig.Rooms[4].IconId := 19;
ApiConfig.Rooms[4].SortDefault := 4;

(* Ručne zvolené ukážkové stavové hodnoty obývačky. *)
ApiState.Rooms[1].RoomId := 1;
ApiState.Rooms[1].Temperature := 22.5;
ApiState.Rooms[1].Humidity := 45.0;
ApiState.Rooms[1].Presence := TRUE;
ApiState.Rooms[1].DayPhase := API_DAY_PHASE_DAY;
ApiState.Rooms[1].CategoryMask := DWORD#16#00000007;
ApiState.Rooms[1].AlarmLevel := API_ALARM_OK;
ApiState.Rooms[1].Online := TRUE;

(* Ručne zvolené ukážkové stavové hodnoty kuchyne. *)
ApiState.Rooms[2].RoomId := 2;
ApiState.Rooms[2].Temperature := 23.0;
ApiState.Rooms[2].Humidity := 48.0;
ApiState.Rooms[2].Presence := FALSE;
ApiState.Rooms[2].DayPhase := API_DAY_PHASE_DUSK;
ApiState.Rooms[2].CategoryMask := DWORD#16#00000003;
ApiState.Rooms[2].AlarmLevel := API_ALARM_WARNING;
ApiState.Rooms[2].Online := TRUE;

(* Ručne zvolené ukážkové stavové hodnoty spálne. *)
ApiState.Rooms[3].RoomId := 3;
ApiState.Rooms[3].Temperature := 21.8;
ApiState.Rooms[3].Humidity := 42.0;
ApiState.Rooms[3].Presence := TRUE;
ApiState.Rooms[3].DayPhase := API_DAY_PHASE_NIGHT;
ApiState.Rooms[3].CategoryMask := DWORD#16#00000001;
ApiState.Rooms[3].AlarmLevel := API_ALARM_OK;
ApiState.Rooms[3].Online := TRUE;

(* Ručne zvolené ukážkové stavové hodnoty terasy. *)
ApiState.Rooms[4].RoomId := 4;
ApiState.Rooms[4].Temperature := 18.4;
ApiState.Rooms[4].Humidity := 58.0;
ApiState.Rooms[4].Presence := FALSE;
ApiState.Rooms[4].DayPhase := API_DAY_PHASE_DAWN;
ApiState.Rooms[4].CategoryMask := DWORD#16#00000004;
ApiState.Rooms[4].AlarmLevel := API_ALARM_ALARM;
ApiState.Rooms[4].Online := FALSE;

(* Tieňové kópie sa zosúladia so snapshotmi, aby štart nevytvoril falošný diff. ENG *)
FOR i := 1 TO C_MAX_ROOMS DO
    ApiConfigShadow[i] := ApiConfig.Rooms[i];
    ApiStateShadow[i] := ApiState.Rooms[i];
END_FOR;

(* Počiatočné verejné informácie a prvý prázdny výsledok príkazu. *)
ApiInfo.ApiVersion := C_API_VERSION;
ApiInfo.ConfigRevision := 1;
ApiInfo.StateRevision := 1;
ApiInfo.MaxRooms := C_MAX_ROOMS;
ApiInfo.LastCommandResult.ClientId := '';
ApiInfo.LastCommandResult.RequestId := 0;
ApiInfo.LastCommandResult.Result := API_RESULT_NONE;
ApiInfo.LastCommandResult.Message := 'Ziadny prikaz';
ApiInfo.LastCommandResult.ConfigRevision := 1;
ApiInfo.LastCommandResult.StateRevision := 1;

(* Pri prvom pripojení musí klient načítať celý konfiguračný snapshot. ENG *)
ApiClearConfigDiff(ApiConfigDiff);
ApiConfigDiff.Valid := TRUE;
ApiConfigDiff.FromRevision := 0;
ApiConfigDiff.ToRevision := 1;
ApiConfigDiff.FullRequired := TRUE;

(* Pri prvom pripojení musí klient načítať celý stavový snapshot. ENG *)
ApiClearStateDiff(ApiStateDiff);
ApiStateDiff.Valid := TRUE;
ApiStateDiff.FromRevision := 0;
ApiStateDiff.ToRevision := 1;
ApiStateDiff.FullRequired := TRUE;

(* Bezpečný počiatočný stav príkazového handshake kanála. ENG *)
ApiCommandRoom.ClientId := '';
ApiCommandRoom.RequestId := 0;
ApiCommandRoom.Action := API_ACTION_NONE;
ApiCommandRoom.RoomId := 0;
ApiCommandRoom.SourceRoomId := 0;
ApiCommandRoom.Name := '';
ApiCommandRoom.ProjectName := '';
ApiCommandExecute := FALSE;
ApiCommandBusy := FALSE;
ApiCommandFinished := FALSE;
ApiCommandResult := ApiInfo.LastCommandResult;

(* Bezpečný počiatočný stav synchronizačného a testovacieho kanála. *)
ApiSyncExecute := FALSE;
ApiSyncBusy := FALSE;
ApiSyncFinished := FALSE;
ApiTestStateExecute := FALSE;
ApiTestStateBusy := FALSE;
ApiTestStateFinished := FALSE;

(* Vynulovanie hláv histórií a pamäte posledného príkazu. *)
ApiConfigHistoryHead := 0;
ApiStateHistoryHead := 0;
ApiLastCommandClientId := '';
ApiLastCommandRequestId := 0;
ApiLastStoredResult := ApiInfo.LastCommandResult;

(* Príznak sa nastaví až po úplnom dokončení celej inicializácie. *)
ApiInitialized := TRUE;
ApiPilotInit := TRUE;
END_FUNCTION

(* ---- 08_COMMAND_ENGINE.ST ---- *)
(* Spracovanie príkazov ADD / DELETE / COPY / SET pre miestnosti. ENG *)

(* Spracuje najviac jeden príkaz, iba ak klient nastavil ApiCommandExecute. *)
FUNCTION ApiProcessRoomCommand : BOOL
VAR
    i             : USINT;     (* Index pri prechode poľom miestností. *)
    configSlot    : USINT;     (* Nájdená alebo voľná pozícia cieľovej konfigurácie. ENG *)
    stateSlot     : USINT;     (* Nájdená alebo voľná pozícia cieľového stavu. ENG *)
    sourceCfgSlot : USINT;     (* Pozícia zdrojovej konfigurácie pri kopírovaní. ENG *)
    sourceStSlot  : USINT;     (* Pozícia zdrojového stavu pri kopírovaní. ENG *)
    maxSort       : UINT;      (* Najvyššie použité predvolené poradie pri pridávaní. ENG *)
    sourceSort    : UINT;      (* Predvolené poradie zdroja pri vkladaní jeho kópie. ENG *)
    deletedSort   : UINT;      (* Predvolené poradie uvoľnené odstránenou miestnosťou. ENG *)
    resultCode    : USINT;     (* Pracovný návratový kód API_RESULT_*. ENG *)
    resultMessage : STRING[80]; (* Pracovný slovenský text výsledku. *)
    executeChange : BOOL;      (* TRUE iba vtedy, keď sa snapshot skutočne zmenil. ENG *)
END_VAR

(* Bez spúšťacieho príznaku funkcia okamžite skončí bez vedľajších účinkov. *)
ApiProcessRoomCommand := FALSE;
IF NOT ApiCommandExecute THEN
    RETURN;
END_IF;

(* Začiatok dvojfázového handshake: príkaz je prevzatý na spracovanie. ENG *)
ApiProcessRoomCommand := TRUE;
ApiCommandBusy := TRUE;
ApiCommandFinished := FALSE;

(* Presné zopakovanie posledného ClientId + RequestId je idempotentné. ENG *)
IF (ApiCommandRoom.ClientId = ApiLastCommandClientId) AND
   (ApiCommandRoom.RequestId = ApiLastCommandRequestId) AND
   (ApiCommandRoom.RequestId <> 0) THEN

    ApiCommandResult := ApiLastStoredResult;
    ApiInfo.LastCommandResult := ApiLastStoredResult;

ELSE
    (* Predvolené hodnoty pre nový, ešte nespracovaný príkaz. *)
    resultCode := API_RESULT_OK;
    resultMessage := 'OK';
    executeChange := FALSE;

    (* Spoločná kontrola povinných identifikátorov transportu. *)
    IF (ApiCommandRoom.ClientId = '') OR (ApiCommandRoom.RequestId = 0) THEN
        resultCode := API_RESULT_INVALID_ARGUMENT;
        resultMessage := 'Neplatny ClientId alebo RequestId';
    ELSE
        (* Rozdelenie spracovania podľa verejného číselného kódu Action. ENG *)
        CASE ApiCommandRoom.Action OF

            API_ACTION_ADD_ROOM:
                (* ADD: overí cieľ, nájde voľné sloty a vytvorí konfiguráciu aj stav. ENG *)
                IF (ApiCommandRoom.RoomId = 0) OR (ApiCommandRoom.Name = '') THEN
                    resultCode := API_RESULT_INVALID_ARGUMENT;
                    resultMessage := 'Neplatne ID alebo nazov';
                ELSIF ApiFindConfigSlot(ApiCommandRoom.RoomId) <> 0 THEN
                    resultCode := API_RESULT_ALREADY_EXISTS;
                    resultMessage := 'RoomId uz existuje';
                ELSE
                    configSlot := ApiFindFreeConfigSlot();
                    stateSlot := ApiFindFreeStateSlot();
                    IF (configSlot = 0) OR (stateSlot = 0) THEN
                        resultCode := API_RESULT_NO_FREE_SLOT;
                        resultMessage := 'Nie je volny slot';
                    ELSE
                        (* Nová miestnosť sa zaradí za najvyššie existujúce SortDefault. ENG *)
                        maxSort := 0;
                        FOR i := 1 TO C_MAX_ROOMS DO
                            IF ApiConfig.Rooms[i].Used AND
                               (ApiConfig.Rooms[i].SortDefault > maxSort) THEN
                                maxSort := ApiConfig.Rooms[i].SortDefault;
                            END_IF;
                        END_FOR;

                        (* Vytvorenie cieľovej konfigurácie z údajov klienta a predvolenej ikony. *)
                        ApiClearRoomConfig(ApiConfig.Rooms[configSlot]);
                        ApiConfig.Rooms[configSlot].Used := TRUE;
                        ApiConfig.Rooms[configSlot].RoomId := ApiCommandRoom.RoomId;
                        ApiConfig.Rooms[configSlot].Name := ApiCommandRoom.Name;
                        ApiConfig.Rooms[configSlot].ProjectName := ApiCommandRoom.ProjectName;
                        ApiConfig.Rooms[configSlot].IconId := API_DEFAULT_ICON_ID;
                        ApiConfig.Rooms[configSlot].SortDefault := maxSort + 1;

                        (* Vytvorenie samostatného stavového záznamu s testovacími hodnotami. *)
                        ApiClearRoomState(ApiState.Rooms[stateSlot]);
                        ApiState.Rooms[stateSlot].RoomId := ApiCommandRoom.RoomId;
                        ApiState.Rooms[stateSlot].Temperature := API_DEFAULT_TEMPERATURE;
                        ApiState.Rooms[stateSlot].Humidity := API_DEFAULT_HUMIDITY;
                        ApiState.Rooms[stateSlot].Presence := FALSE;
                        ApiState.Rooms[stateSlot].DayPhase := API_DAY_PHASE_DAY;
                        ApiState.Rooms[stateSlot].CategoryMask := DWORD#16#00000000;
                        ApiState.Rooms[stateSlot].AlarmLevel := API_ALARM_OK;
                        ApiState.Rooms[stateSlot].Online := TRUE;

                        executeChange := TRUE;
                        resultMessage := 'Miestnost pridana';
                    END_IF;
                END_IF;

            API_ACTION_DELETE_ROOM:
                (* DELETE: konfigurácia aj stav musia existovať, potom sa oba sloty vyčistia. ENG *)
                configSlot := ApiFindConfigSlot(ApiCommandRoom.RoomId);
                stateSlot := ApiFindStateSlot(ApiCommandRoom.RoomId);
                IF (configSlot = 0) OR (stateSlot = 0) THEN
                    resultCode := API_RESULT_NOT_FOUND;
                    resultMessage := 'Miestnost nenajdena';
                ELSE
                    (* Uložené poradie sa použije na zhutnenie hodnôt po zmazaní. *)
                    deletedSort := ApiConfig.Rooms[configSlot].SortDefault;
                    ApiClearRoomConfig(ApiConfig.Rooms[configSlot]);
                    ApiClearRoomState(ApiState.Rooms[stateSlot]);

                    (* Miestnosti za odstránenou pozíciou sa posunú o jedno miesto dopredu. *)
                    FOR i := 1 TO C_MAX_ROOMS DO
                        IF ApiConfig.Rooms[i].Used AND
                           (ApiConfig.Rooms[i].SortDefault > deletedSort) THEN
                            ApiConfig.Rooms[i].SortDefault :=
                                ApiConfig.Rooms[i].SortDefault - 1;
                        END_IF;
                    END_FOR;

                    executeChange := TRUE;
                    resultMessage := 'Miestnost zmazana';
                END_IF;

            API_ACTION_COPY_ROOM:
                (* COPY: najprv sa overí zdroj aj jedinečnosť cieľového RoomId. ENG *)
                sourceCfgSlot := ApiFindConfigSlot(ApiCommandRoom.SourceRoomId);
                sourceStSlot := ApiFindStateSlot(ApiCommandRoom.SourceRoomId);
                IF (ApiCommandRoom.RoomId = 0) OR
                   (ApiCommandRoom.RoomId = ApiCommandRoom.SourceRoomId) THEN
                    resultCode := API_RESULT_INVALID_ARGUMENT;
                    resultMessage := 'Neplatne cielove RoomId';
                ELSIF (sourceCfgSlot = 0) OR (sourceStSlot = 0) THEN
                    resultCode := API_RESULT_NOT_FOUND;
                    resultMessage := 'Zdrojova miestnost nenajdena';
                ELSIF ApiFindConfigSlot(ApiCommandRoom.RoomId) <> 0 THEN
                    resultCode := API_RESULT_ALREADY_EXISTS;
                    resultMessage := 'Cielove RoomId uz existuje';
                ELSE
                    configSlot := ApiFindFreeConfigSlot();
                    stateSlot := ApiFindFreeStateSlot();
                    IF (configSlot = 0) OR (stateSlot = 0) THEN
                        resultCode := API_RESULT_NO_FREE_SLOT;
                        resultMessage := 'Nie je volny slot';
                    ELSE
                        (* Pre kópiu sa uvoľní poradie hneď za zdrojovou miestnosťou. *)
                        sourceSort := ApiConfig.Rooms[sourceCfgSlot].SortDefault;
                        FOR i := 1 TO C_MAX_ROOMS DO
                            IF ApiConfig.Rooms[i].Used AND
                               (ApiConfig.Rooms[i].SortDefault > sourceSort) THEN
                                ApiConfig.Rooms[i].SortDefault :=
                                    ApiConfig.Rooms[i].SortDefault + 1;
                            END_IF;
                        END_FOR;

                        (* Konfigurácia sa kopíruje celá; klient môže voliteľne prepísať názvy. *)
                        ApiConfig.Rooms[configSlot] := ApiConfig.Rooms[sourceCfgSlot];
                        ApiConfig.Rooms[configSlot].RoomId := ApiCommandRoom.RoomId;
                        ApiConfig.Rooms[configSlot].SortDefault := sourceSort + 1;
                        IF ApiCommandRoom.Name <> '' THEN
                            ApiConfig.Rooms[configSlot].Name := ApiCommandRoom.Name;
                        END_IF;
                        IF ApiCommandRoom.ProjectName <> '' THEN
                            ApiConfig.Rooms[configSlot].ProjectName := ApiCommandRoom.ProjectName;
                        END_IF;

                        (* Pilot kopíruje aj ručne nastavený stav, ale priradí nové RoomId. ENG *)
                        ApiState.Rooms[stateSlot] := ApiState.Rooms[sourceStSlot];
                        ApiState.Rooms[stateSlot].RoomId := ApiCommandRoom.RoomId;

                        executeChange := TRUE;
                        resultMessage := 'Miestnost skopirovana';
                    END_IF;
                END_IF;

            API_ACTION_SET_ROOM_DATA:
                (* SET: v pilote mení iba hlavný a doplnkový názov miestnosti. ENG *)
                configSlot := ApiFindConfigSlot(ApiCommandRoom.RoomId);
                IF configSlot = 0 THEN
                    resultCode := API_RESULT_NOT_FOUND;
                    resultMessage := 'Miestnost nenajdena';
                ELSIF ApiCommandRoom.Name = '' THEN
                    resultCode := API_RESULT_INVALID_ARGUMENT;
                    resultMessage := 'Nazov nesmie byt prazdny';
                ELSE
                    ApiConfig.Rooms[configSlot].Name := ApiCommandRoom.Name;
                    ApiConfig.Rooms[configSlot].ProjectName := ApiCommandRoom.ProjectName;
                    executeChange := TRUE;
                    resultMessage := 'Udaje miestnosti nastavene';
                END_IF;

            ELSE
                (* Neznámy číselný kód Action sa odmietne bez zmeny dát. ENG *)
                resultCode := API_RESULT_UNSUPPORTED_ACTION;
                resultMessage := 'Nepodporovana akcia';
        END_CASE;
    END_IF;

    (* Úspešná dátová zmena vytvorí nové revízie a príslušné diff rámce. ENG *)
    IF executeChange AND (resultCode = API_RESULT_OK) THEN
        ApiCaptureConfigChanges();
        ApiCaptureStateChanges();
    END_IF;

    (* Výsledok nesie identitu požiadavky aj revízie platné po jej spracovaní. *)
    ApiCommandResult.ClientId := ApiCommandRoom.ClientId;
    ApiCommandResult.RequestId := ApiCommandRoom.RequestId;
    ApiCommandResult.Result := resultCode;
    ApiCommandResult.Message := resultMessage;
    ApiCommandResult.ConfigRevision := ApiInfo.ConfigRevision;
    ApiCommandResult.StateRevision := ApiInfo.StateRevision;

    (* Uloženie výsledku pre ApiInfo a idempotentné opakovanie poslednej požiadavky. *)
    ApiInfo.LastCommandResult := ApiCommandResult;
    ApiLastCommandClientId := ApiCommandRoom.ClientId;
    ApiLastCommandRequestId := ApiCommandRoom.RequestId;
    ApiLastStoredResult := ApiCommandResult;
END_IF;

(* Ukončenie handshake: PLC zruší Execute, uvoľní Busy a nastaví Finished. ENG *)
ApiCommandExecute := FALSE;
ApiCommandBusy := FALSE;
ApiCommandFinished := TRUE;
END_FUNCTION

(* ---- 09_STATE_TEST.ST ---- *)
(* Ručný validovaný zápis testovacieho stavu; nie je pripojené žiadne reálne IO. *)

(* Spracuje najviac jednu testovaciu požiadavku po nastavení ApiTestStateExecute. *)
FUNCTION ApiProcessTestState : BOOL
VAR
    configSlot    : USINT;      (* Pozícia konfigurácie cieľovej miestnosti. ENG *)
    stateSlot     : USINT;      (* Pozícia stavového záznamu cieľovej miestnosti. ENG *)
    resultCode    : USINT;      (* Pracovný návratový kód API_RESULT_*. ENG *)
    resultMessage : STRING[80]; (* Pracovný slovenský text výsledku. *)
END_VAR

(* Bez spúšťacieho príznaku funkcia skončí bez vedľajších účinkov. *)
ApiProcessTestState := FALSE;
IF NOT ApiTestStateExecute THEN
    RETURN;
END_IF;

(* Prevzatie požiadavky a nastavenie predvoleného úspešného výsledku. *)
ApiProcessTestState := TRUE;
ApiTestStateBusy := TRUE;
ApiTestStateFinished := FALSE;
resultCode := API_RESULT_OK;
resultMessage := 'Testovaci stav nastaveny';

(* Miestnosť musí existovať súčasne v konfigurácii aj v stavovom snapshote. *)
configSlot := ApiFindConfigSlot(ApiTestStateRequest.RoomId);
stateSlot := ApiFindStateSlot(ApiTestStateRequest.RoomId);

(* Validácia identity požiadavky, existencie miestnosti a povolených rozsahov. *)
IF (ApiTestStateRequest.ClientId = '') OR
   (ApiTestStateRequest.RequestId = 0) THEN
    resultCode := API_RESULT_INVALID_ARGUMENT;
    resultMessage := 'Neplatny ClientId alebo RequestId';
ELSIF (configSlot = 0) OR (stateSlot = 0) THEN
    resultCode := API_RESULT_NOT_FOUND;
    resultMessage := 'Miestnost nenajdena';
ELSIF (ApiTestStateRequest.Temperature < -50.0) OR
      (ApiTestStateRequest.Temperature > 100.0) OR
      (ApiTestStateRequest.Humidity < 0.0) OR
      (ApiTestStateRequest.Humidity > 100.0) OR
      (ApiTestStateRequest.AlarmLevel > API_ALARM_ALARM) OR
      (NOT ApiValidDayPhase(ApiTestStateRequest.DayPhase)) THEN
    resultCode := API_RESULT_INVALID_ARGUMENT;
    resultMessage := 'Neplatna testovacia hodnota';
ELSE
    (* Platné hodnoty sa zapíšu iba do dynamického stavu, nie do konfigurácie. *)
    ApiState.Rooms[stateSlot].Temperature := ApiTestStateRequest.Temperature;
    ApiState.Rooms[stateSlot].Humidity := ApiTestStateRequest.Humidity;
    ApiState.Rooms[stateSlot].Presence := ApiTestStateRequest.Presence;
    ApiState.Rooms[stateSlot].DayPhase := ApiTestStateRequest.DayPhase;
    ApiState.Rooms[stateSlot].CategoryMask := ApiTestStateRequest.CategoryMask;
    ApiState.Rooms[stateSlot].AlarmLevel := ApiTestStateRequest.AlarmLevel;
    ApiState.Rooms[stateSlot].Online := ApiTestStateRequest.Online;
    ApiCaptureStateChanges();
END_IF;

(* Výsledok obsahuje identitu požiadavky a revízie platné po spracovaní. *)
ApiTestStateResult.ClientId := ApiTestStateRequest.ClientId;
ApiTestStateResult.RequestId := ApiTestStateRequest.RequestId;
ApiTestStateResult.Result := resultCode;
ApiTestStateResult.Message := resultMessage;
ApiTestStateResult.ConfigRevision := ApiInfo.ConfigRevision;
ApiTestStateResult.StateRevision := ApiInfo.StateRevision;

(* Ukončenie testovacieho handshake kanála. ENG *)
ApiTestStateExecute := FALSE;
ApiTestStateBusy := FALSE;
ApiTestStateFinished := TRUE;
END_FUNCTION

(* ---- 10_SYNC_ENGINE.ST ---- *)
(* Obnova cache: vráti jeden ďalší uchovaný rámec alebo vyžiada celý snapshot. ENG *)

(* Pripraví odpoveď na jednu synchronizačnú požiadavku klienta. *)
FUNCTION ApiProcessSyncRequest : BOOL
VAR
    i           : USINT; (* Index pri prehľadávaní kruhových histórií diffov. *)
    foundConfig : BOOL;  (* TRUE po nájdení platnej odpovede pre konfiguráciu. ENG *)
    foundState  : BOOL;  (* TRUE po nájdení platnej odpovede pre stav. ENG *)
END_VAR

(* Bez spúšťacieho príznaku funkcia skončí bez vedľajších účinkov. *)
ApiProcessSyncRequest := FALSE;
IF NOT ApiSyncExecute THEN
    RETURN;
END_IF;

(* Prevzatie synchronizačnej požiadavky na spracovanie. *)
ApiProcessSyncRequest := TRUE;
ApiSyncBusy := TRUE;
ApiSyncFinished := FALSE;

(* Identita odpovede sa vždy kopíruje z aktuálnej požiadavky klienta. *)
ApiSyncResponse.ClientId := ApiSyncRequest.ClientId;
ApiSyncResponse.RequestId := ApiSyncRequest.RequestId;
ApiSyncResponse.Result := API_RESULT_OK;
ApiSyncResponse.Message := 'Synchronizacia pripravena';

(* Pred hľadaním sa vyčistia oba výstupné rámce a pomocné príznaky. *)
ApiClearConfigDiff(ApiSyncResponse.ConfigDiff);
ApiClearStateDiff(ApiSyncResponse.StateDiff);
foundConfig := FALSE;
foundState := FALSE;

(* Neplatná identita sa oznámi v Result; režimy diffov sa napriek tomu určia deterministicky. ENG *)
IF (ApiSyncRequest.ClientId = '') OR (ApiSyncRequest.RequestId = 0) THEN
    ApiSyncResponse.Result := API_RESULT_INVALID_ARGUMENT;
    ApiSyncResponse.Message := 'Neplatny ClientId alebo RequestId';
END_IF;

(* Konfiguračná vetva: CURRENT, jeden nadväzujúci DIFF alebo FULL_REQUIRED. ENG *)
IF ApiSyncRequest.ConfigFromRevision = ApiInfo.ConfigRevision THEN
    ApiSyncResponse.ConfigMode := API_SYNC_CURRENT;
    ApiSyncResponse.ConfigDiff.Valid := TRUE;
    ApiSyncResponse.ConfigDiff.FromRevision := ApiInfo.ConfigRevision;
    ApiSyncResponse.ConfigDiff.ToRevision := ApiInfo.ConfigRevision;
    foundConfig := TRUE;
ELSE
    FOR i := 1 TO C_DIFF_HISTORY_DEPTH DO
        IF ApiConfigDiffHistory[i].Valid AND
           (ApiConfigDiffHistory[i].FromRevision =
            ApiSyncRequest.ConfigFromRevision) THEN
            ApiSyncResponse.ConfigDiff := ApiConfigDiffHistory[i];
            ApiSyncResponse.ConfigMode := API_SYNC_DIFF;
            foundConfig := TRUE;
            EXIT;
        END_IF;
    END_FOR;
END_IF;

(* Ak požadovaná revízia už nie je v histórii, klient musí načítať celý snapshot. *)
IF NOT foundConfig THEN
    ApiSyncResponse.ConfigMode := API_SYNC_FULL_REQUIRED;
    ApiSyncResponse.ConfigDiff.Valid := TRUE;
    ApiSyncResponse.ConfigDiff.FromRevision := ApiSyncRequest.ConfigFromRevision;
    ApiSyncResponse.ConfigDiff.ToRevision := ApiInfo.ConfigRevision;
    ApiSyncResponse.ConfigDiff.FullRequired := TRUE;
END_IF;

(* Stavová vetva: CURRENT, jeden nadväzujúci DIFF alebo FULL_REQUIRED. ENG *)
IF ApiSyncRequest.StateFromRevision = ApiInfo.StateRevision THEN
    ApiSyncResponse.StateMode := API_SYNC_CURRENT;
    ApiSyncResponse.StateDiff.Valid := TRUE;
    ApiSyncResponse.StateDiff.FromRevision := ApiInfo.StateRevision;
    ApiSyncResponse.StateDiff.ToRevision := ApiInfo.StateRevision;
    foundState := TRUE;
ELSE
    FOR i := 1 TO C_DIFF_HISTORY_DEPTH DO
        IF ApiStateDiffHistory[i].Valid AND
           (ApiStateDiffHistory[i].FromRevision =
            ApiSyncRequest.StateFromRevision) THEN
            ApiSyncResponse.StateDiff := ApiStateDiffHistory[i];
            ApiSyncResponse.StateMode := API_SYNC_DIFF;
            foundState := TRUE;
            EXIT;
        END_IF;
    END_FOR;
END_IF;

(* Ak požadovaná stavová revízia nie je v histórii, klient načíta celý snapshot. *)
IF NOT foundState THEN
    ApiSyncResponse.StateMode := API_SYNC_FULL_REQUIRED;
    ApiSyncResponse.StateDiff.Valid := TRUE;
    ApiSyncResponse.StateDiff.FromRevision := ApiSyncRequest.StateFromRevision;
    ApiSyncResponse.StateDiff.ToRevision := ApiInfo.StateRevision;
    ApiSyncResponse.StateDiff.FullRequired := TRUE;
END_IF;

(* Ukončenie synchronizačného handshake kanála. ENG *)
ApiSyncExecute := FALSE;
ApiSyncBusy := FALSE;
ApiSyncFinished := TRUE;
END_FUNCTION

(* ---- prgMain.ST ---- *)
(* Hlavn� cyklick� program ROOM_API_PILOT vykon�van� PLC. *)
PROGRAM prgMain
VAR
    (* Program z�merne nepotrebuje �iadne lok�lne premenn�. *)
END_VAR

(* Jednorazov� inicializ�cia; po prvom �spe�nom cykle u� d�ta nemen�. *)
ApiPilotInit();

IF ApiInitialized THEN
	SizeApiHeder 	:= SIZEOF(NH_API_DIFF_HEAD);
	SizeStructRoom := SIZEOF(T_ROOM_STATE);
	SizeApiVars		:= SIZEOF(ApiVarsPublic);
	Ptr_T_ROOM_STATE_Dest^ := Ptr_T_ROOM_STATE_Src^;

    (* Najprv sa spracuj poiadavky, ktor mu zmeni konfigurciu alebo stav. *)
    ApiProcessRoomCommand();
    ApiProcessTestState();

    (* Zachyt aj run zmeny vykonan cez okno Watch v Mosaic. ENG *)
    ApiCaptureConfigChanges();
    ApiCaptureStateChanges();

    (* Synchroniz�cia sa spracuje a� po zachyten� v�etk�ch zmien dan�ho cyklu. *)
    ApiProcessSyncRequest();
END_IF;
END_PROGRAM
